TYPE ST_FORCE_REF : FB_FORCE_REF;
END_TYPE

(* stored: Version 1.1.0.1, ProductVersion 3.1.4024.15
   DUT ST_FORCE_REF: Id {fbdf3630-3c09-4691-a73b-fb34872b1bb6} *)
